DATA_BLOCK "DB_Mando"
{ S7_Optimized_Access := 'TRUE' }
VERSION : 0.1
NON_RETAIN
"FB_Mando_Motor"

BEGIN

END_DATA_BLOCK

